RoboDK station: Simulacion_brazorobotico.rdk

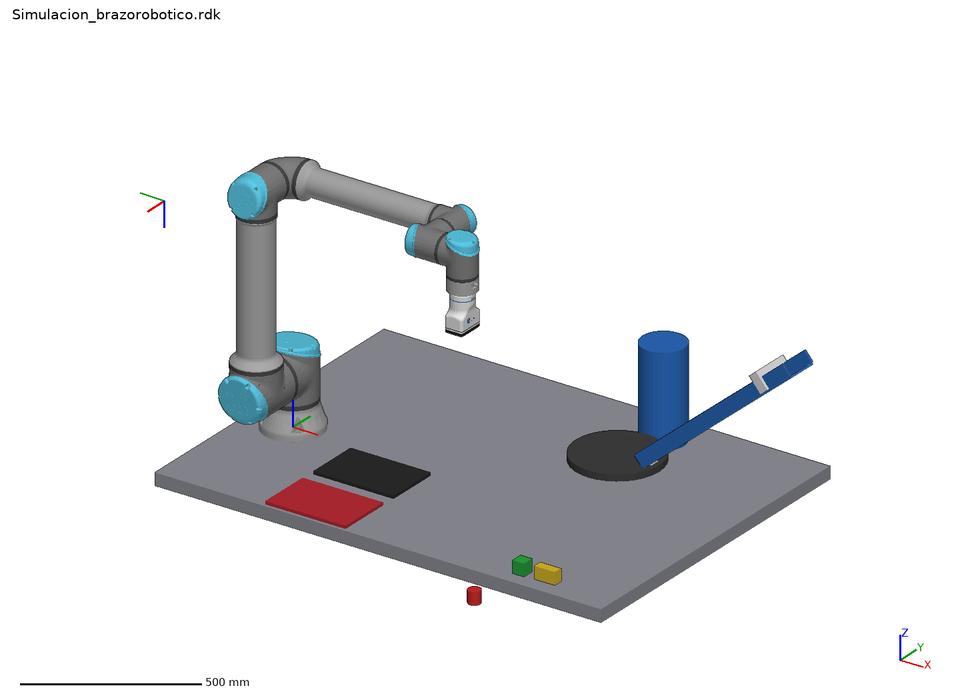
[picture v0: the station drawn from its stored meshes, robots at their saved joint values, targets as dots, program paths as lines]
Station Nueva Estación 1 (saved by RoboDK 6.0.7). Poses are relative to the parent item; angles as X-Y-Z fixed-axis rotations.
  - frame UR10e Base at (0, 0, 0) mm
    - robot UR10e: 6 axes, payload 10 kg, reach 1300 mm, repeatability 0.05 mm, weight 28.9 kg
        modified DH rows (alpha deg, a mm, theta deg, d mm): 0, 0, 0, 180.7; 90, 0, 180, 0; 0, 612.6, 0, 0; 0, 571.335, 0, 174.15; -90, 0, 0, 119.85; 90, 0, 180, 116.55
        joint limits [-360, -360, -360, -360, -360, -360] to [360, 360, 360, 360, 360, 360]; home [0, -90, -90, 0, 90, 0]; saved at [0, -90, -90, -90, 90, 0]
      - robot OnRobot 2FG7 Gripper: 1 axes
          joint limits [0] to [55]; home [0]; saved at [0]
      - frame Pinza at (0, 1000, 0) mm
  - Python program Prog1 (listed below)
  - frame Celda at (0, 0, 0) mm
    - object Mesa at (600, 100, -20) mm, size 1500 x 1100 x 40 mm, geometry from Mesa.stl
    - object Bandeja_Roja at (350, -350, 5) mm, size 270 x 180 x 10 mm, geometry from Bandeja_Roja.stl
    - object Bandeja_Negra at (350, -120, 5) mm, size 270 x 180 x 10 mm, geometry from Bandeja_Negra.stl
    - object Reductor at (880, 300, 15) mm, size 100 x 100 x 30 mm, geometry from Reductor.stl
    - object Plato at (880, 300, 40) mm, size 280 x 280 x 20 mm, geometry from Plato.stl
    - object Marcador_Plato at (990, 300, 51.5) mm, size 30 x 30 x 3 mm, geometry from Marcador_Plato.stl
    - object Sistema_Vision at (880, 520, 150) mm, size 140 x 140 x 300 mm, geometry from Sistema_Vision.stl
    - object Rampa_Fondo at (1250.89, 300, 266.61) mm, rotated rx 0 ry -40 rz 0 deg, size 650 x 100 x 6 mm, geometry from Rampa_Fondo.stl
    - object Rampa_Pared1 at (1236.11, 353, 284.23) mm, rotated rx 0 ry -40 rz 0 deg, size 650 x 6 x 40 mm, geometry from Rampa_Pared1.stl
    - object Rampa_Pared2 at (1236.11, 247, 284.23) mm, rotated rx 0 ry -40 rz 0 deg, size 650 x 6 x 40 mm, geometry from Rampa_Pared2.stl
    - object Dosificador at (1398.21, 300, 433.3) mm, rotated rx 0 ry -40 rz 0 deg, size 30 x 130 x 60 mm, geometry from Dosificador.stl
    - object Pieza_cilindro at (1145, -765, 110) mm, rotated rx -180 ry 0 rz -90 deg, size 40 x 40 x 40 mm, geometry from Pieza_cilindro.stl
    - object Pieza_cubo at (1145, -535, 110) mm, rotated rx 180 ry 0 rz -90 deg, size 40 x 40 x 40 mm, geometry from Pieza_cubo.stl
    - object Pieza_prisma at (1230, -535, 110) mm, rotated rx -180 ry 0 rz -90 deg, size 30 x 70 x 40 mm, geometry from Pieza_prisma.stl

--- Python program Prog1 ---
import os, math, tempfile, time
from robodk.robolink import *
from robodk.robomath import *

RDK = Robolink()
TMP = tempfile.mkdtemp()

def msg(t, popup=False):
    print(t)
    RDK.ShowMessage(str(t), popup)

# ====== MEDIDAS (mm), RELATIVAS A LA BASE DEL ROBOT. AJUSTA CON TU CELDA ======
Z_TCP       = 150                 # distancia brida -> puntas de los dedos
C_PLATO     = (880, 300)          # centro del plato giratorio
PLATO_TOP   = 50                  # altura de la cara superior del plato
P_RAMPA     = transl(1000, 300, 60) * roty(math.radians(-40))  # extremo bajo de la rampa
LARGO_RAMPA = 650
SLOT0, PASO = 400, 50             # posiciones de espera de las piezas en la rampa
ENTRADA     = (950, 300)          # donde cae la pieza sobre el plato
PICK        = transl(880, 370, 70) * rotx(math.pi)   # pieza sobre el plato tras girar 90 deg
BANDEJA_ROJA  = (350, -350)
BANDEJA_NEGRA = (350, -120)
HOME = [0, -90, -90, -90, 90, 0]
# nombre, color RGBA, bandeja destino
TIPOS = [('cilindro', [0.9, 0.1, 0.1, 1], 'roja'),
         ('cubo',     [0.1, 0.7, 0.2, 1], 'negra'),
         ('prisma',   [0.95, 0.8, 0.1, 1], 'negra')]
# =================================================================================

NOMBRES = ['Celda', 'Mesa', 'Bandeja_Roja', 'Bandeja_Negra', 'Reductor', 'Plato',
           'Marcador_Plato', 'Sistema_Vision', 'Rampa_Fondo', 'Rampa_Pared1',
           'Rampa_Pared2', 'Dosificador', 'TCP_Pinza'] + ['Pieza_' + t[0] for t in TIPOS]

# ---------- Geometria (STL) ----------
def _stl(nombre, tris):
    ruta = os.path.join(TMP, nombre + '.stl')
    with open(ruta, 'w') as f:
        f.write('solid %s\n' % nombre)
        for t in tris:
            f.write('facet normal 0 0 0\nouter loop\n')
            for v in t:
                f.write('vertex %f %f %f\n' % tuple(v))
            f.write('endloop\nendfacet\n')
        f.write('endsolid\n')
    return ruta

def caja(sx, sy, sz):
    x, y, z = sx/2, sy/2, sz/2
    v = [(-x,-y,-z),(x,-y,-z),(x,y,-z),(-x,y,-z),(-x,-y,z),(x,-y,z),(x,y,z),(-x,y,z)]
    c = [(0,2,1),(0,3,2),(4,5,6),(4,6,7),(0,1,5),(0,5,4),
         (1,2,6),(1,6,5),(2,3,7),(2,7,6),(3,0,4),(3,4,7)]
    return [[v[i] for i in f] for f in c]

def cilindro(r, h, n=32):
    t, z = [], h/2
    for i in range(n):
        a0, a1 = 2*math.pi*i/n, 2*math.pi*(i+1)/n
        p0 = (r*math.cos(a0), r*math.sin(a0)); p1 = (r*math.cos(a1), r*math.sin(a1))
        t.append([(p0[0],p0[1],-z),(p1[0],p1[1],-z),(p1[0],p1[1],z)])
        t.append([(p0[0],p0[1],-z),(p1[0],p1[1],z),(p0[0],p0[1],z)])
        t.append([(0,0,z),(p0[0],p0[1],z),(p1[0],p1[1],z)])
        t.append([(0,0,-z),(p1[0],p1[1],-z),(p0[0],p0[1],-z)])
    return t

def crear(nombre, tris, pose, color, padre):
    it = RDK.AddFile(_stl(nombre, tris), padre)
    it.setName(nombre)
    it.setPose(pose)          # pose local respecto al marco 'Celda'
    it.setColor(color)
    return it

# ---------- Robot y base ----------
def buscar_robot():
    for it in RDK.ItemList(ITEM_TYPE_ROBOT):
        try:
            if len(it.Joints().list()) == 6:
                return it
        except Exception:
            pass
    r = RDK.Item('UR10e', ITEM_TYPE_ROBOT)
    if not r.Valid():
        raise Exception("No se encontro el robot UR10e (6 ejes) en la estacion")
    return r

def obtener_base(robot):
    padre = robot.Parent()
    if padre.Valid() and padre.Type() == ITEM_TYPE_FRAME:
        return padre.PoseAbs()
    msg('AVISO: el robot no esta dentro de un marco de base; uso el origen de la estacion.')
    return eye(4)

def limpiar():
    for n in NOMBRES:
        for _ in range(5):
            it = RDK.Item(n)
            if not it.Valid():
                break
            it.Delete()

# ---------- Construccion de la celda ----------
def construir(celda):
    gris, blanco, azul = [0.6,0.6,0.65,1], [0.95,0.95,0.95,1], [0.1,0.4,0.8,1]
    cx, cy = C_PLATO
    crear('Mesa', caja(1500, 1100, 40), transl(600, 100, -20), gris, celda)
    crear('Bandeja_Roja',  caja(270, 180, 10), transl(*BANDEJA_ROJA, 5),  [0.8,0.1,0.15,1], celda)
    crear('Bandeja_Negra', caja(270, 180, 10), transl(*BANDEJA_NEGRA, 5), [0.1,0.1,0.1,1], celda)
    crear('Reductor', caja(100, 100, 30), transl(cx, cy, 15), blanco, celda)
    crear('Plato', cilindro(140, 20), transl(cx, cy, 40), [0.2,0.2,0.2,1], celda)
    crear('Marcador_Plato', caja(30, 30, 3), transl(cx+110, cy, PLATO_TOP+1.5), [1,1,1,1], celda)
    crear('Sistema_Vision', cilindro(70, 300), transl(cx, cy+220, 150), azul, celda)
    L = LARGO_RAMPA
    crear('Rampa_Fondo',  caja(L, 100, 6),  P_RAMPA*transl(L/2, 0, -3),  azul, celda)
    crear('Rampa_Pared1', caja(L, 6, 40),   P_RAMPA*transl(L/2, 53, 20), azul, celda)
    crear('Rampa_Pared2', caja(L, 6, 40),   P_RAMPA*transl(L/2, -53, 20), azul, celda)
    crear('Dosificador',  caja(30, 130, 60), P_RAMPA*transl(545, 0, 30), blanco, celda)
    formas = {'cilindro': cilindro(20, 40), 'cubo': caja(40, 40, 40), 'prisma': caja(30, 70, 40)}
    for i, (nombre, color, _) in enumerate(TIPOS):
        crear('Pieza_' + nombre, formas[nombre], P_RAMPA*transl(SLOT0 + PASO*i, 0, 20), color, celda)

# ---------- Utilidades de simulacion ----------
def girar(items, grados, pasos=30):
    cx, cy = C_PLATO
    for i in range(1, pasos + 1):
        R = transl(cx, cy, 0) * rotz(math.radians(grados*i/pasos)) * transl(-cx, -cy, 0)
        for it, p0 in items:
            it.setPose(R * p0)
        RDK.Render(True)
        time.sleep(0.03)

def deslizar(pieza, x0, x1=20, pasos=40):
    for i in range(pasos + 1):
        x = x0 + (x1 - x0) * i / pasos
        pieza.setPose(P_RAMPA * transl(x, 0, 20))
        RDK.Render(True)
        time.sleep(0.02)

def huecos(c):
    return [transl(c[0]+dx, c[1]+dy, 30) * rotx(math.pi) for dy in (-45, 45) for dx in (-85, 0, 85)]

def mover(robot, tipo, destino, paso):
    msg(paso)
    try:
        if tipo == 'J':
            robot.MoveJ(destino)
        else:
            robot.MoveL(destino)
    except Exception as e:
        if tipo == 'L':
            try:
                robot.MoveJ(destino)      # plan B: movimiento articular
                return
            except Exception:
                pass
        raise Exception('Fallo el movimiento "%s": %s' % (paso, e))

# ---------- Programa principal ----------
def main():
    msg('1/6 Preparando simulacion')
    RDK.setRunMode(RUNMODE_SIMULATE)
    RDK.setSimulationSpeed(1)
    robot = buscar_robot()
    base = obtener_base(robot)

    msg('2/6 Limpiando celda anterior')
    limpiar()
    celda = RDK.AddFrame('Celda')
    celda.setPose(base)

    msg('3/6 Construyendo celda')
    construir(celda)

    msg('4/6 Configurando robot')
    robot.setPoseTool(transl(0, 0, Z_TCP))
    robot.setSpeed(500)
    robot.setSpeedJoints(90)
    robot.setJoints(HOME)

    marcador = RDK.Item('Marcador_Plato')
    contador = {'roja': 0, 'negra': 0}
    bandejas = {'roja': huecos(BANDEJA_ROJA), 'negra': huecos(BANDEJA_NEGRA)}

    msg('5/6 Piezas en la rampa; el robot va a HOME')
    mover(robot, 'J', HOME, 'Robot a HOME')

    msg('6/6 Inicio del ciclo de clasificacion')
    for i, (nombre, _, destino) in enumerate(TIPOS):
        pieza = RDK.Item('Pieza_' + nombre)
        msg('Pieza %s: baja por la rampa' % nombre)
        deslizar(pieza, SLOT0 + PASO*i)
        pieza.setPose(transl(ENTRADA[0], ENTRADA[1], PLATO_TOP + 20))
        msg('Pieza %s: el plato gira hacia la vision' % nombre)
        girar([(pieza, pieza.Pose()), (marcador, marcador.Pose())], 90)
        msg('Vision: pieza detectada -> %s | destino: bandeja %s' % (nombre, destino))
        time.sleep(1)

        mover(robot, 'J', PICK * transl(0, 0, -120), 'Aproximar a ' + nombre)
        mover(robot, 'L', PICK, 'Bajar a tomar ' + nombre)
        pieza.setParentStatic(robot)                      # agarrar
        mover(robot, 'L', PICK * transl(0, 0, -120), 'Subir con ' + nombre)

        hueco = bandejas[destino][contador[destino]]
        contador[destino] += 1
        mover(robot, 'J', hueco * transl(0, 0, -120), 'Ir a la bandeja ' + destino)
        mover(robot, 'L', hueco, 'Bajar a dejar ' + nombre)
        pieza.setParentStatic(celda)                      # soltar
        mover(robot, 'L', hueco * transl(0, 0, -120), 'Subir de la bandeja')
        mover(robot, 'J', HOME, 'Volver a HOME')
        girar([(marcador, marcador.Pose())], -90)          # el plato vuelve

    msg('Simulacion terminada: 3 piezas clasificadas', True)

try:
    main()
except Exception as e:
    RDK.ShowMessage('ERROR: ' + str(e), True)
    raise
